// Mitsubishi GX Works2 project: AVRInfacomV4   PLC: FX3G

TYPE CutCard : STRUCT
  Lenth : DINT;
  Qnt : DINT;
END_STRUCT END_TYPE

// global labels: _io
VAR_GLOBAL
  DI_Avar1 AT X000 : BOOL;  (* Сигнал аварии автомата Сети 1: 0 — авария по логике ПЛК *)
  DI_Line1IsOff AT X001 : BOOL;  (* Обратная связь автомата Сети 1: 1 — разомкнут *)
  DI_Avar2 AT X002 : BOOL;  (* Сигнал аварии автомата Сети 2: 0 — авария по логике ПЛК *)
  DI_Line2IsOff AT X003 : BOOL;  (* Обратная связь автомата Сети 2: 1 — разомкнут *)
  DI_AvarGenerator AT X004 : BOOL;  (* Сигнал аварии автомата генератора: 0 — авария по логике ПЛК *)
  DI_GeneratorIsOff AT X005 : BOOL;  (* Обратная связь автомата генератора: 1 — разомкнут *)
  DI_AvarSection AT X006 : BOOL;  (* Резерв: вход аварии секционного автомата *)
  DI_SectionIsOff AT X007 : BOOL;  (* Резерв: обратная связь секционного автомата *)
  DI_RKF1 AT X010 : BOOL;  (* Сигнал РКФ Сети 1: 1 — параметры источника в норме *)
  DI_RKF2 AT X011 : BOOL;  (* Сигнал РКФ Сети 2: 1 — параметры источника в норме *)
  DI_RKF3 AT X012 : BOOL;  (* Сигнал РКФ генератора: 1 — параметры источника в норме *)
  DI_Avarkontrol AT X013 : BOOL;  (* Вспомогательный контакт общего автомата питания приводов после ИБП; 1 — норма по логике ПЛК *)
  DO_On1 AT Y000 : BOOL;  (* Выход включения автомата Сети 1 *)
  DO_Off1 AT Y001 : BOOL;  (* Выход отключения автомата Сети 1 *)
  DO_On2 AT Y002 : BOOL;  (* Выход включения автомата Сети 2 *)
  DO_Off2 AT Y003 : BOOL;  (* Выход отключения автомата Сети 2 *)
  DO_OnGenerator AT Y004 : BOOL;  (* Выход включения автомата генератора *)
  DO_OffGenerator AT Y005 : BOOL;  (* Выход отключения автомата генератора *)
  DO_OnSection AT Y006 : BOOL;  (* Резерв: выход включения секционного автомата *)
  DO_OffSection AT Y007 : BOOL;  (* Резерв: выход отключения секционного автомата *)
  DO_StartGenerator AT Y010 : BOOL;  (* Расчётный выход запроса запуска генератора: 0 — запрос; запуск выполняет внешняя автоматика *)
END_VAR

// global labels: _gvl
VAR_GLOBAL
  gxAvto AT M400 : BOOL;  (* Режим АВР: 1 — автоматический, 0 — ручной *)
  gxOn1 AT M100 : BOOL;  (* Тогл включения автомата Сети 1 на панели; ПЛК может сбросить *)
  gxOff1 AT M101 : BOOL;  (* Ручная команда отключения автомата Сети 1 *)
  gxOn2 AT M102 : BOOL;  (* Тогл включения автомата Сети 2 на панели; ПЛК может сбросить *)
  gxOff2 AT M103 : BOOL;  (* Ручная команда отключения автомата Сети 2 *)
  gxOnGenerator AT M104 : BOOL;  (* Тогл включения автомата генератора на панели; ПЛК может сбросить *)
  gxOffGenerator AT M105 : BOOL;  (* Ручная команда отключения автомата генератора *)
  gxOnSection AT M106 : BOOL;  (* Резерв: команда включения секционного автомата *)
  gxOffSection AT M107 : BOOL;  (* Резерв: команда отключения секционного автомата *)
  gxStartGenerator AT M108 : BOOL;  (* Ручной запрос запуска генератора в программе; фактический запуск внешний *)
  gxIsAlarm AT M150 : BOOL;  (* Общий признак наличия аварий *)
  gxVVAOff AT M401 : BOOL;  (* Защёлкнутый общий признак неисправности ВА; выбором источника не используется *)
  gxProblemVVA1 AT M110 : BOOL;  (* Защёлкнутый отказ включения или неожиданное размыкание автомата Сети 1 *)
  gxProblemVVA2 AT M111 : BOOL;  (* Защёлкнутый отказ включения или неожиданное размыкание автомата Сети 2 *)
  gxProblemVVAgen AT M112 : BOOL;  (* Защёлкнутый отказ включения или неожиданное размыкание автомата генератора *)
  clTimeGenerator AT D1000 : INT;  (* Уставка таймера импульса запуска генератора, с *)
  clTimeRKF1 AT D1001 : INT;  (* Задержка подтверждения готовности Сети 1, с *)
  clTimeRKF2 AT D1002 : INT;  (* Задержка подтверждения готовности Сети 2, с *)
  clTimeRKF3 AT D1003 : INT;  (* Задержка подтверждения готовности генератора, с *)
  clStartgenerator AT D1004 : INT;  (* Тайм-аут подтверждения напряжения после запроса запуска генератора, с *)
  clTimeBackAuto AT D1005 : INT;  (* Уставка задержки возврата в AUTO, с; логика закомментирована *)
  VVALine1 : VVA;  (* Экземпляр блока управления автоматом Сети 1 *)
  VVALine2 : VVA;  (* Экземпляр блока управления автоматом Сети 2 *)
  VVAGen : VVA;  (* Экземпляр блока управления автоматом генератора *)
  VVASec : VVA;  (* Экземпляр блока секционного автомата; в управлении не вызывается *)
END_VAR

// task Task_init (event M8002, interval 0, priority 1): PRG_INIT
// task Task_Main (event TRUE, interval 0, priority 31): PGN_MAIN
// task Task_Process (event TRUE, interval 0, priority 31): PRG_PROCESS
// user libraries (not included): AlarmManger128, Modbusv16, TimeControl, Utils

PROGRAM PGN_MAIN
VAR
  fbAmBlock : AM_IS_BLOCK;  (* Проверка блокирующих аварий; вызов закомментирован *)
  fbAmalarm : AM_HAS_ALARMS;  (* Проверка наличия аварий для общего признака gxIsAlarm *)
  fbTPStartGen : TP;  (* Таймер импульса запроса запуска генератора *)
  xGenerator : BOOL;  (* Внутренний запрос запуска генератора *)
  xDrivePower : BOOL;  (* Разрешение по X13; принудительно снято в первом скане RUN *)
  xAllOff : BOOL;  (* Все три автомата по обратной связи разомкнуты *)
  xAutoWasOn : BOOL;  (* Режим AUTO в предыдущем скане для обнаружения смены режима *)
  xManualOn1 : BOOL;  (* Фронт команды включения автомата Сети 1 с панели *)
  xManualOn2 : BOOL;  (* Фронт команды включения автомата Сети 2 с панели *)
  xManualOnGen : BOOL;  (* Фронт команды включения автомата генератора с панели *)
  xSetOn1 : BOOL;  (* Удерживаемая заявка на включение автомата Сети 1, не импульс *)
  xSetOn2 : BOOL;  (* Удерживаемая заявка на включение автомата Сети 2, не импульс *)
  xSetOnGen : BOOL;  (* Удерживаемая заявка на включение автомата генератора, не импульс *)
  iStep : INT;  (* Шаг АВР: 0 — пуск, 10 — ожидание или ручной режим, 20 — выбор, 30/40/50 — источники *)
END_VAR
(* fbAmBlock(iProcessNum := 1, iSeverity := AM_ERROR, Q := gxIsAlarm); *)
fbAmalarm(
    iProcessNum := 0,
    iSeverity := 0,
    Q := gxIsAlarm
);

(* Предполагается, что при исправном общем питании на X13 высокий уровень. M8002
   принудительно выполняет сброс в первом цикле после перехода в RUN, даже если X13 уже активен. *)
xDrivePower := DI_Avarkontrol AND NOT M8002;
(* Нормально замкнутые контакты положения дают TRUE при отключённом выключателе. *)
xAllOff := DI_Line1IsOff AND DI_Line2IsOff AND DI_GeneratorIsOff;
(* В каждом цикле ПЛК отслеживать передние фронты ручных команд включения. Команда,
   поданная во время запрета, не запоминается: после снятия запрета нужно нажать кнопку снова. *)
xManualOn1 := MEP(gxOn1);
xManualOn2 := MEP(gxOn2);
xManualOnGen := MEP(gxOnGenerator);

IF xAutoWasOn <> gxAvto THEN
    IF NOT gxAvto THEN
        (* Переход из автоматического режима в ручной: взять фактические положения, а не ожидающие команды.
           Для включённого выключателя сохранить запрос на включённое положение, даже если автоматика запрашивала отключение.
           Для отключённого выключателя оставить запрос снятым, отменив ожидающие попытки включения. *)
        xSetOn1 := NOT DI_Line1IsOff;
        xSetOn2 := NOT DI_Line2IsOff;
        xSetOnGen := NOT DI_GeneratorIsOff;
    ELSE
        (* При переходе в автоматический режим перед выбором источника отменить невыполненные ручные запросы на включение. *)
        xSetOn1 := xSetOn1 AND NOT DI_Line1IsOff;
        xSetOn2 := xSetOn2 AND NOT DI_Line2IsOff;
        xSetOnGen := xSetOnGen AND NOT DI_GeneratorIsOff;
    END_IF;
    IF iStep <> 0 THEN
        iStep := 10; (* Вернуться к ручному управлению или выбору источника, а не к шагу прежнего источника. *)
    END_IF;
END_IF;

(* Источник доступен, только если реле контроля фаз и аппаратный вход контроля аварии
   показывают норму, а у выключателя нет зафиксированной тревоги или неисправности. *)
M1 := DI_RKF1 AND DI_Avar1 AND NOT VVALine1.xError AND NOT gxProblemVVA1;
M2 := DI_RKF2 AND DI_Avar2 AND NOT VVALine2.xError AND NOT gxProblemVVA2;
M3 := DI_RKF3 AND DI_AvarGenerator AND NOT VVAGen.xError AND NOT gxProblemVVAgen;

OUT_T(M1, TC1, SEC_TO_TIMER100(clTimeRKF1));
OUT_T(M2, TC2, SEC_TO_TIMER100(clTimeRKF2));
OUT_T(M3, TC3, SEC_TO_TIMER100(clTimeRKF3));

(* TC30 отсчитывает время при наличии сигнала исправности питания приводов: 100 × 100 мс = 10 с.
   Пропадание сигнала X13 сбрасывает таймер. Во время ожидания на шаге 0 все прежние запросы снимаются. *)
OUT_T(xDrivePower, TC30, K100);
IF NOT xDrivePower OR NOT TS30 THEN
    iStep := 0;
END_IF;

(* Перед новым автоматическим запросом на включение выдержать паузу: все три сигнала
   отключённого положения должны непрерывно оставаться активными, а запросов на включение быть не должно.
   После отмены запроса не переносить отсчитанное время на другой источник. Номинальная выдержка при K11 — 1,1 с. *)
OUT_T(
    gxAvto
    AND xDrivePower
    AND xAllOff
    AND NOT (xSetOn1 OR xSetOn2 OR xSetOnGen),
    TC32,
    K11
);

(* Возврат в автоматический режим
OUT_T(gxVVAOff, TC31, SEC_TO_TIMER100(clTimeBackAuto));
IF TS31 THEN
	gxVVAOff := FALSE;
END_IF;
 *)

CASE iStep OF
    0: (* Ожидание питания приводов, взвода пружин и отключённого положения выключателей. *)
        xGenerator := FALSE;
        gxStartGenerator := FALSE;
        xSetOn1 := FALSE;
        xSetOn2 := FALSE;
        xSetOnGen := FALSE;
        (* Выйти из пускового шага только после выдержки времени, когда все три выключателя отключены. *)
        MOV(
            xDrivePower
            AND TS30
            AND xAllOff,
            10,
            iStep
        );

    10: (* Ожидание или ручное управление. *)
        IF gxAvto THEN
            iStep := 20;
            gxStartGenerator := FALSE;
        ELSIF NOT xAutoWasOn AND NOT M2002 AND xAllOff AND NOT (xSetOn1 OR xSetOn2 OR xSetOnGen) THEN
            (* В предыдущем цикле должен быть ручной режим. Не должно быть квитирования
               или действующего запроса; все выключатели должны быть отключены. Цепочка ELSIF
               принимает не более одного запроса на включение: сначала ввод 1, затем ввод 2, затем генератор. *)
            IF xManualOn1 AND M1 AND NOT gxOff1 THEN
                xSetOn1 := TRUE;
            ELSIF xManualOn2 AND M2 AND NOT gxOff2 THEN
                xSetOn2 := TRUE;
            ELSIF xManualOnGen AND M3 AND NOT gxOffGenerator THEN
                xSetOnGen := TRUE;
            END_IF;
        END_IF;
        IF NOT gxAvto THEN
            (* Команда отключения, потеря готовности источника или включение другого выключателя
               отменяют соответствующий ручной запрос и его повторные попытки. *)
            RST(
                gxOff1
                OR NOT DI_Line2IsOff
                OR NOT DI_GeneratorIsOff
                OR NOT M1,
                xSetOn1
            );
            RST(
                gxOff2
                OR NOT DI_Line1IsOff
                OR NOT DI_GeneratorIsOff
                OR NOT M2,
                xSetOn2
            );
            RST(
                gxOffGenerator
                OR NOT DI_Line1IsOff
                OR NOT DI_Line2IsOff
                OR NOT M3,
                xSetOnGen
            );
        END_IF;
        xGenerator := gxStartGenerator;

    20: (* Выбрать первый доступный источник после выдержки времени по сигналу реле контроля фаз. *)
        MOV(TS1, 30, iStep);
        MOV(
            TS2
            AND NOT TS1,
            40,
            iStep
        );
        MOV(
            NOT TS1
            AND NOT TS2
            AND TS3,
            50,
            iStep
        );
        (* Сохранить запрос на включение только для выбранного источника, остальные снять. *)
        xSetOn1 := xSetOn1 AND iStep = 30;
        xSetOn2 := xSetOn2 AND iStep = 40;
        xSetOnGen := xSetOnGen AND iStep = 50;
        xGenerator := NOT TS1 AND NOT TS2;

    30: (* Ввод 1. Такая же блокировка действует на шагах 40 и 50. *)
        (* Снять запросы на включение двух других выключателей, чтобы их блоки могли подать команды отключения. *)
        xSetOn2 := FALSE;
        xSetOnGen := FALSE;
        MOV(
            NOT TS1 (* Ввод 1 больше не готов. *)
            OR NOT M1, (* Ввод 1 больше не удовлетворяет условиям доступности, проверяемым без задержки. *)
            10,
            iStep
        );
        (* Выдерживать паузу только перед новым запросом. Сохранять действующий запрос,
           когда его выключатель включается и сбрасывает TC32 или когда VVA ещё выполняет повторные попытки. *)
        xSetOn1 := DI_GeneratorIsOff
            AND DI_Line2IsOff
            AND iStep = 30
            AND (xSetOn1 OR (xAllOff AND TS32));

    40: (* Ввод 2: перед запросом на включение дождаться отключения выключателей ввода 1 и генератора. *)
        xSetOn1 := FALSE;
        xSetOnGen := FALSE;
        MOV(
            NOT TS2 (* Ввод 2 больше не готов. *)
            OR NOT M2, (* Ввод 2 больше не удовлетворяет условиям доступности, проверяемым без задержки. *)
            10,
            iStep
        );
        xSetOn2 := DI_GeneratorIsOff
            AND DI_Line1IsOff
            AND iStep = 40
            AND (xSetOn2 OR (xAllOff AND TS32));

    50: (* Генератор: дождаться отключения выключателей обоих сетевых вводов. Вернуться к выбору источника,
           если один из сетевых вводов снова готов или генератор больше недоступен. *)
        xSetOn2 := FALSE;
        xSetOn1 := FALSE;
        MOV(
            NOT TS3 (* Готовность по напряжению генератора больше не подтверждается. *)
            OR NOT M3 (* Генератор больше не удовлетворяет условиям доступности, проверяемым без задержки. *)
            OR TS1 OR TS2, (* Готов хотя бы один сетевой ввод. *)
            10,
            iStep
        );
        xGenerator := TRUE;
        xSetOnGen := DI_Line1IsOff
            AND DI_Line2IsOff
            AND iStep = 50
            AND (xSetOnGen OR (xAllOff AND TS32));
ELSE (* Недопустимый номер шага: снять запросы и вернуться к пусковому шагу. *)
    iStep := 0;
    xSetOn1 := FALSE;
    xSetOn2 := FALSE;
    xSetOnGen := FALSE;
END_CASE;
xAutoWasOn := gxAvto; (* Запомнить режим, чтобы обнаружить его смену в следующем цикле ПЛК. *)

fbTPStartGen(
    IN := xGenerator,
    PT := SEC_TO_TIME(clTimeGenerator)
);
DO_StartGenerator := NOT (xGenerator OR fbTPStartGen.Q);

(* Вызывать блок каждого выключателя в каждом цикле, в том числе при пуске, чтобы таймеры
   и выходы обновлялись даже без запроса на включение. Для IsOn инвертировать сигнал отключённого положения. *)
VVALine1(
    SetOn := xSetOn1,
    IsOn := NOT DI_Line1IsOff,
    xDrivePower := xDrivePower,
    ResetAlarm := M2002,
    Vkl := DO_On1,
    Otkl := DO_Off1
);
VVALine2(
    SetOn := xSetOn2,
    IsOn := NOT DI_Line2IsOff,
    xDrivePower := xDrivePower,
    ResetAlarm := M2002,
    Vkl := DO_On2,
    Otkl := DO_Off2
);
VVAGen(
    SetOn := xSetOnGen,
    IsOn := NOT DI_GeneratorIsOff,
    xDrivePower := xDrivePower,
    ResetAlarm := M2002,
    Vkl := DO_OnGenerator,
    Otkl := DO_OffGenerator
);

(* В ручном режиме сбросить переключатель «Вкл.» на панели оператора только при отключённом выключателе:
   если нет действующего запроса или блок только что сообщил об исчерпании попыток включения.
   Не сбрасывать переключатель в паузах между попытками и после успешного включения. *)
IF NOT gxAvto THEN
    RST(
        DI_Line1IsOff
        AND (NOT xSetOn1 OR VVALine1.xVklFailed),
        gxOn1
    );
    RST(
        DI_Line2IsOff
        AND (NOT xSetOn2 OR VVALine2.xVklFailed),
        gxOn2
    );
    RST(
        DI_GeneratorIsOff
        AND (NOT xSetOnGen OR VVAGen.xVklFailed),
        gxOnGenerator
    );
END_IF;

(* Зафиксировать исчерпание попыток включения или неожиданное отключение. Со следующего цикла
   проверка доступности исключает этот выключатель, пока неисправность не будет сброшена. *)
SET(
    VVALine1.xVklFailed
    OR VVALine1.xUnexpectedOff,
    gxProblemVVA1
);
SET(
    VVALine2.xVklFailed
    OR VVALine2.xUnexpectedOff,
    gxProblemVVA2
);
SET(
    VVAGen.xVklFailed
    OR VVAGen.xUnexpectedOff,
    gxProblemVVAgen
);
SET(
    gxProblemVVA1
    OR gxProblemVVA2
    OR gxProblemVVAgen,
    gxVVAOff
);
END_PROGRAM

PROGRAM PRG_INIT
VAR
  fbAmInit : AM_INIT;  (* Регистрация аварий при инициализации *)
END_VAR
AM_D_START := 3000;

VVALine1.AlarmNum := 1;
VVALine2.AlarmNum := 2;
VVAGen.AlarmNum := 3;
VVASec.AlarmNum := 4;

(* Ошибка UPS *)
fbAmInit(iNum := 0, iSeverity := 3, iProcess := 1, xLatch := 0, xBuzzer := 0, xLock := 0);
(* Ошибка ВА Сеть 1 *)
fbAmInit(iNum := 1 , xLatch := 1, xLock := 0 );
(* Ошибка ВА Сеть 2 *)
fbAmInit(iNum := 2 , xLatch := 1, xLock := 0 );
(* Ошибка ВА Генератор *)
fbAmInit(iNum := 3 , xLatch := 1, xLock := 0 );
(* Ошибка ВА Секционный *)
fbAmInit(iNum := 4 , xLatch := 1, xLock := 0);
(* Отказ вкл ВА Сеть 1 *)
fbAmInit(iNum := 5, xLatch := 0, xLock := 0);
(* Отказ выкл ВА Сеть 1 *)
fbAmInit(iNum := 6 , xLatch := 0, xLock := 0 );
(* Отказ вкл ВА Сеть 2 *)
fbAmInit(iNum := 7 , xLatch := 0, xLock := 0 );
(* Отказ выкл ВА Сеть 2 *)
fbAmInit(iNum := 8 , xLatch := 0, xLock := 0 );
(* Отказ вкл ВА Генератор *)
fbAmInit(iNum := 9 , xLatch := 0, xLock := 0);
(* Отказ выкл ВА Генератор *)
fbAmInit(iNum := 10, xLatch := 0, xLock := 0);
(* Отказ вкл ВА Секционный *)
fbAmInit(iNum := 11 , xLatch := 0, xLock := 0 );
(* Отказ выкл ВА Секционный *)
fbAmInit(iNum := 12 , xLatch := 0, xLock := 0 );
(* Отказ запуска генератора *)
fbAmInit(iNum := 13 , xLatch := 1, xLock := 0 );
(* Данные не заполнены *)
fbAmInit(iNum := 14 , xLatch := 0, xLock := 1);
END_PROGRAM

PROGRAM PRG_PROCESS
VAR
  fbAmSet : AM_SET;  (* Передача состояния аварии в менеджер по её номеру *)
  fbAmReset : AM_RST;  (* Квитирование аварий по команде M2002 *)
  fbAMEvents : AM_EVENT;  (* Регистрация событий в журнале *)
  fbTOFResetProblems : TOF;  (* Таймер отложенного сброса неисправностей; вызов закомментирован *)
  xNodata : BOOL;  (* Хотя бы одна проверяемая временная уставка равна нулю *)
  xMBInit : BOOL;  (* Результат вызова инициализации Modbus RTU; не признак связи *)
  PortSettings : DWORD;  (* Настройки порта Modbus RTU: 38400 бод, без чётности, 1 стоп-бит *)
END_VAR
fbAmReset(IN := M2002);

IF M2002 THEN
	gxProblemVVA1 := FALSE;
	gxProblemVVA2 := FALSE;
	gxProblemVVAgen := FALSE;
END_IF;

PortSettings := MB_PORT_SETTINGS(MB_PARITY_NONE, MB_STOPBIT_1, MB_BPS_38400);
xMBInit := MB_SLAVE_INIT_PORT2(TRUE, 20, PortSettings);

(* Тревоги *)
OUT_T(NOT DI_Avarkontrol, TC24, 10);
fbAmSet(iNum := 0, xState := TS24);
(* Для тревог 1–3 запустить таймер на 500 мс в одном из двух случаев:
   - X13 и TC30 подтверждают восстановление питания приводов, но вход контроля отдельного выключателя имеет низкий уровень;
   - PRG_MAIN уже зафиксировала исчерпание попыток включения или неожиданное отключение.
   Зафиксированная неисправность выключателя отображается даже при пропадании общего питания. *)
OUT_T(
    (DI_Avarkontrol AND TS30 AND NOT DI_Avar1)
    OR gxProblemVVA1,
    TC21,
    5
);
fbAmSet(iNum := 1, xState := TS21);
OUT_T(
    (DI_Avarkontrol AND TS30 AND NOT DI_Avar2)
    OR gxProblemVVA2,
    TC22,
    5
);
fbAmSet(iNum := 2, xState := TS22);
OUT_T(
    (DI_Avarkontrol AND TS30 AND NOT DI_AvarGenerator)
    OR gxProblemVVAgen,
    TC23,
    5
);
fbAmSet(iNum := 3, xState := TS23);
fbAmSet(iNum := 4, xState := FALSE);
OUT_T(DO_On1 AND DI_Line1IsOff, TC11, 10);
fbAmSet(iNum := 5, xState := TS11);
OUT_T(DO_Off1 AND NOT DI_Line1IsOff, TC12, 10);
fbAmSet(iNum := 6, xState := TS12);
OUT_T(DO_On2 AND DI_Line2IsOff, TC13, 10);
fbAmSet(iNum := 7, xState := TS13);
OUT_T(DO_Off2 AND NOT DI_Line2IsOff, TC14, 10);
fbAmSet(iNum := 8, xState := TS14);
OUT_T(DO_Ongenerator AND DI_GeneratorIsOff, TC15, 10);
fbAmSet(iNum := 9, xState := TS15);
OUT_T(DO_OffGenerator AND NOT DI_GeneratorIsOff, TC16, 10);
fbAmSet(iNum := 10, xState := TS16);
(* Здесь нет проверки включения секционного выключателя: прежняя проверка тоже записывала
   состояние тревоги 1 и могла перезаписать состояние тревоги ввода 1 в том же цикле ПЛК. *)
OUT_T(DO_OffSection AND NOT DI_SectionIsOff, TC18, 10);
fbAmSet(iNum := 12, xState := TS18);
OUT_T(NOT DO_StartGenerator AND NOT DI_RKF3, TC19, SEC_TO_TIMER100(clStartgenerator));
fbAmSet(iNum := 13, xState := TS19);

xNodata := (
	clStartgenerator = 0
	OR clTimeGenerator = 0
	OR clTimeRKF1 = 0
	OR clTimeRKF2 = 0
	OR clTimeRKF3 = 0
);
fbAmSet(iNum := 14, xState := xNodata);

fbAMEvents(EventNum := 0, EventState := DI_RKF1);
fbAMEvents(EventNum := 1, EventState := NOT DI_RKF1);
fbAMEvents(EventNum := 2, EventState := DI_RKF2);
fbAMEvents(EventNum := 3, EventState := NOT DI_RKF2);
fbAMEvents(EventNum := 4, EventState := DI_RKF3);
fbAMEvents(EventNum := 5, EventState := NOT DI_RKF3);
fbAMEvents(EventNum := 6, EventState := DO_On1);
fbAMEvents(EventNum := 7, EventState := DO_Off1);
fbAMEvents(EventNum := 8, EventState := DO_On2);
fbAMEvents(EventNum := 9, EventState := DO_Off2);
fbAMEvents(EventNum := 10, EventState := DO_Ongenerator);
fbAMEvents(EventNum := 11, EventState := DO_Offgenerator);
fbAMEvents(EventNum := 12, EventState := DO_OnSection);
fbAMEvents(EventNum := 13, EventState := DO_OffSection);
fbAMEvents(EventNum := 14, EventState := NOT DO_StartGenerator);
fbAMEvents(EventNum := 15, EventState := DO_StartGenerator);
fbAMEvents(EventNum := 16, EventState := gxAvto);
fbAMEvents(EventNum := 17, EventState := NOT gxAvto);
fbAMEvents(EventNum := 18, EventState := TS1);
fbAMEvents(EventNum := 19, EventState := TS2);
fbAMEvents(EventNum := 20, EventState := TS3);

(*
fbTOFResetProblems(IN:= MEP(gxProblemVVA1) OR MEP(gxProblemVVA2) OR MEP(gxProblemVVAgen), PT:= SEC_TO_TIME(1800));
IF M2002 OR fbTOFResetProblems.Q THEN
	gxProblemVVA1 := FALSE;
	gxProblemVVA2 := FALSE;
	gxProblemVVAgen := FALSE;
END_IF;
 *)
END_PROGRAM

FUNCTION_BLOCK VVA
VAR_INPUT
  SetOn : BOOL;  (* Запрошенное положение: 1 — замкнуть или удерживать замкнутым *)
  xDrivePower : BOOL;  (* Разрешение работы привода от ПЛК по состоянию общего питания *)
  IsOn : BOOL;  (* Текущее положение по обратной связи: 1 — автомат замкнут *)
  ResetAlarm : BOOL;  (* Команда квитирования аварии *)
  AlarmNum : INT;  (* Номер аварии этого автомата в менеджере аварий *)
END_VAR
VAR_OUTPUT
  Vkl : BOOL;  (* Импульс включения автомата *)
  Otkl : BOOL;  (* Импульс отключения автомата *)
  xError : BOOL;  (* Защёлкнутая авария автомата; запрещает включение *)
  xVklFailed : BOOL;  (* Отказ включения: импульс на один скан после трёх неудачных попыток *)
  xUnexpectedOff : BOOL;  (* Подтверждённое неожиданное размыкание при действующей заявке на включение *)
END_VAR
VAR
  fbAmIsOn : AM_ORISON;  (* Чтение состояния аварии по номеру AlarmNum *)
  fbBlinkOff : BLINK;  (* Формирование повторных импульсов отключения *)
  fbTONOn : TON;  (* Подтверждение замкнутого положения за 100 мс *)
  fbTONOff : TON;  (* Подтверждение разомкнутого положения за 100 мс *)
  fbVklPulse : TON;  (* Таймер импульса включения на 900 мс *)
  fbVklWait : TON;  (* Пауза 7 с после импульса включения перед повтором или отказом *)
  xTempError : BOOL;  (* Результат чтения аварии в текущем скане; сбрасывается перед вызовом *)
  xWasClosed : BOOL;  (* Память: при текущей заявке уже подтверждалось замкнутое положение *)
  iVklStep : INT;  (* Шаг цикла включения: 0 — ожидание, 10 — импульс, 20 — пауза, 30 — отказ *)
  iVklAttempts : INT;  (* Количество начатых попыток включения для текущей заявки *)
END_VAR
(* SetOn — запрошенное положение, IsOn — фактическое положение.
   Vkl и Otkl — выходы включения и отключения. Блок не меняет режим управления. *)

(* При квитировании сбросить зафиксированную ошибку блока, затем проверить, сохраняется ли её причина.
   Перед вызовом библиотечного блока обнулить временный результат: если Q не будет записан
   в этом цикле ПЛК, значение TRUE из предыдущего цикла не должно снова установить xError. *)
RST(xError AND ResetAlarm, xError);
xTempError := FALSE;
fbAmIsOn(
    iNum := AlarmNum,
    Q := xTempError
);
SET(xTempError, xError); (* Активная тревога снова устанавливает xError даже при квитировании. *)

(* Подтверждать положение только после 100 мс стабильного сигнала обратной связи. *)
fbTONOn(
    IN := IsOn,
    PT := T#100ms
);
fbTONOff(
    IN := NOT IsOn,
    PT := T#100ms
);
(* Каждый таймер сбрасывается вне своего шага. Первый завершает импульс включения;
   второй отсчитывает паузу 7 с для привода после снятия сигнала включения. *)
fbVklPulse(
    IN := iVklStep = 10,
    PT := T#900ms
);
fbVklWait(
    IN := iVklStep = 20,
    PT := T#7s
);

(* Пересчитывать сигналы неисправности в каждом цикле ПЛК. PRG_MAIN фиксирует обнаруженную неисправность. *)
xVklFailed := FALSE;
xUnexpectedOff := FALSE;
IF NOT xDrivePower OR NOT SetOn OR xError THEN
    (* Как только запрос становится недопустимым, снять сигнал включения и отменить повторные попытки. *)
    xWasClosed := FALSE;
    iVklStep := 0;
    iVklAttempts := 0;
ELSIF fbTONOn.Q THEN
    (* Включение подтверждено. Запомнить это до снятия запроса. *)
    xWasClosed := TRUE;
    iVklStep := 0;
    iVklAttempts := 0;
ELSIF xWasClosed THEN
    (* Не считать отключение после подтверждённого включения отказом включения. *)
    xUnexpectedOff := fbTONOff.Q;
ELSE
    CASE iVklStep OF
        0: (* Первая попытка: только при подтверждённом отключении и без активного сигнала квитирования. *)
            IF fbTONOff.Q AND NOT ResetAlarm THEN
                iVklAttempts := 1;
                iVklStep := 10;
            END_IF;
        10: (* Импульс включения: завершить по таймеру или сразу при появлении сигнала IsOn. *)
            IF fbVklPulse.Q OR IsOn THEN
                iVklStep := 20;
            END_IF;
        20: (* Сигнал включения снят. Через 7 с повторить попытку, только если отключённое положение всё ещё подтверждается. *)
            IF fbVklWait.Q AND fbTONOff.Q AND NOT ResetAlarm THEN
                IF iVklAttempts < K3 THEN
                    iVklAttempts := iVklAttempts + K1;
                    iVklStep := 10; (* Возврат на шаг 10 формирует новый передний фронт сигнала включения. *)
                ELSE
                    xVklFailed := TRUE; (* После третьей попытки выдать сигнал отказа на один цикл ПЛК. *)
                    iVklStep := 30;
                END_IF;
            END_IF;
        30: (* После трёх попыток не подавать сигнал включения, пока запрос не снят. *)
            iVklStep := 30;
    ELSE (* При недопустимом номере шага вернуться к ожиданию. *)
        iVklStep := 0;
        iVklAttempts := 0;
    END_CASE;
END_IF;

(* Шаги заменяют fbBlinkOn: на шаге 10 — импульс, на шаге 20 — пауза, затем шаг 10 даёт новый фронт.
   Перед записью выхода в каждом цикле ПЛК заново проверять все условия включения в блоке. *)
Vkl := xDrivePower AND SetOn AND NOT xError AND NOT IsOn AND iVklStep = 10;

(* Отключение не зависит от шагов включения. Отключать замкнутый выключатель, если
   снят запрос на включение или активна тревога. Подавать импульсы до размыкания;
   последнее AND сразу снимает сигнал отключения, если запрос на отключение исчез. *)
Otkl := xDrivePower AND (NOT SetOn OR xError) AND IsOn;
fbBlinkOff(
    IN := Otkl,
    TIMELOW := T#1000ms,
    TIMEHIGH := T#1000ms
);
Otkl := Otkl AND fbBlinkOff.Q;
END_FUNCTION_BLOCK
